// TIA Portal V19 export
// export: Created 2026-10-15T09:44:23.0228615Z, ExportSetting WithDefaults, DisplayName Totally Integrated Automation Portal, DisplayVersion V19, DisplayName TIA Portal Openness, DisplayVersion V19, DisplayName TIA Portal Version Control Interface, DisplayVersion V19, DisplayName STEP 7 Professional, DisplayVersion V19, DisplayName STEP 7 Safety, DisplayVersion V19, DisplayName WinCC Basic/Comfort/Advanced, DisplayVersion V19, DisplayName WinCC Unified, DisplayVersion V19
FUNCTION "ROLL_EncodeSeconds" : Word   // FC5, SCL
{ S7_Optimized_Access := 'TRUE' }
VERSION : 0.1
// stored: AutoNumber true, IsIECCheckEnabled false, SetENOAutomatically false, UDAEnableTagReadback false
   VAR_INPUT
      Seconds : Int;
   END_VAR
BEGIN

   IF (#Seconds < 0) OR (#Seconds > 999) THEN
       #ROLL_EncodeSeconds := W#16#FFFF;
   ELSE
       #ROLL_EncodeSeconds := W#16#2000 OR SHL(IN := INT_TO_WORD(#Seconds / 100), N := 8)
       OR SHL(IN := INT_TO_WORD((#Seconds / 10) MOD 10), N := 4) OR INT_TO_WORD(#Seconds MOD 10);
   END_IF;
END_FUNCTION
